// TIA Portal V20 export
// export: Created 2026-10-21T13:28:37.0680677Z, ExportSetting None, DisplayName Totally Integrated Automation Portal, DisplayVersion V20, DisplayName TIA Portal Openness, DisplayVersion V20, DisplayName TIA Portal Version Control Interface, DisplayVersion V20, DisplayName STEP 7 Professional, DisplayVersion V20, DisplayName STEP 7 Safety, DisplayVersion V20, DisplayName WinCC Basic/Comfort/Advanced, DisplayVersion V20, DisplayName WinCC Unified, DisplayVersion V20
DATA_BLOCK "iDB_M01"   // DB1
AUTHOR : JMellid
FAMILY : Drives
// Al generar este bloque, TIA crea el DB de instancia "iDB_M01" del FB_Motor.
// ==============================================================================
// stored: InstanceOfName FB_Motor, InstanceOfType FB
"FB_Motor"
   // VAR_INPUT
   //    CmdStart : Bool;
   //    CmdStop : Bool;
   //    CmdReset : Bool;
   //    Interlock : Bool;
   //    Feedback : Bool;
   //    FeedbackUsed : Bool;
   //    StartTimeout : Time;
   //    StopTimeout : Time;
   // END_VAR
   // VAR_OUTPUT
   //    Run : Bool;
   //    Running : Bool;
   //    Ready : Bool;
   //    Fault : Bool;
   //    FaultCode : Int;
   // END_VAR
   // VAR
   //    statRunLatch : Bool;
   //    statWasConfirmed : Bool;
   //    statFault : Bool;
   //    statFaultCode : Int;
   //    tonStart { S7_SetPoint := 'True'} : TON_TIME;
   //    tonStop { S7_SetPoint := 'True'} : TON_TIME;
   // END_VAR
BEGIN
END_DATA_BLOCK
